Fanuc KAREL source: kc00018.KL

-- PROVISIONAL review KL for V1013-1; original PC SHA256 7c8a0142ed7e2e78518883b096752f689fe145895729e759ddd1006e534d6e16
-- Incomplete behavior may be omitted. Consult companion uncertainty JSON. Do not deploy.
PROGRAM KC00018
%NOLOCKGROUP
BEGIN
  -- UNRESOLVED_PC offsets 5-63; opcodes 27,22,2A,22,2A,22,22,2A,22,22,22,22,31
  -- UNRESOLVED_PC offsets 68-72; opcodes 7F
END KC00018
